// SIMATIC S7-200 project (STEP 7-Micro/WIN), CPU 224 CN REL 02.01

SYMBOL_TABLE USUARIO1
SF               I0.3     // Sensor de objetos
SII              I0.4     // Sensor inductivo (Metal)
SP               I0.5     // Sensor magnetico (plastico)
SM1              I0.7     // Sensor magnetico extendido 1
SM2              I1.0     // Sensor magnetico extendido 2
SM3              I1.1     // Sensor magnetico extendido 3
SB_2             I1.2     // Pulsador de paro
SB_1             I1.3     // Pulsador de marcha
QS               I1.4     // Zeta de emergencia
SA               I1.5     // Selector de modo
Motor            Q0.0     // Motor
KV1              Q0.4     // Cilindro neumatico 1
KV2              Q0.5     // Cilindro neumatico 2
KV3              Q0.6     // Cilindro neumatico 3
HL1              Q0.7     // Piloto indicador de parada
HL2              Q1.0     // Piloto indicador de marcha
HL3              Q1.1     // Piloto indicador de emergencia
E0               M0.0
E1               M0.1
E2               M0.2
E3               M0.3
E4               M0.4
E5               M0.5
E6               M0.6
E7               M0.7
E8               M1.0
E9               M1.1
EP               M1.2
EM               M1.3
END_CTRL         M1.4     // bit de finalizacion del controlador
C_1              VD100
L_k              VD110
r_k              VD120
e_k              VD130
U_k              VD150
Kp               VD160
END_SYMBOL_TABLE

ORGANIZATION_BLOCK PRINCIPAL:OB1
TITLE=COMENTARIOS DEL PROGRAMA
BEGIN
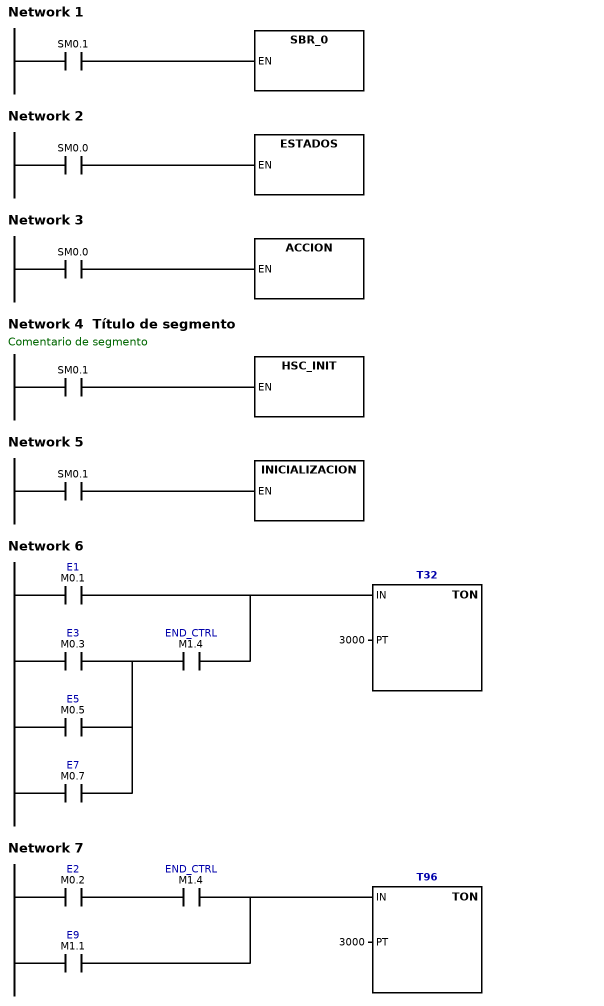
Network 1
LD     SM0.1
CALL   SBR_0:SBR0
Network 2
LD     SM0.0
CALL   ESTADOS:SBR3
Network 3
LD     SM0.0
CALL   ACCION:SBR4
Network 4 // Título de segmento
// Comentario de segmento
LD     SM0.1
CALL   HSC_INIT:SBR1
Network 5
LD     SM0.1
CALL   INICIALIZACION:SBR2
Network 6
LD     E1:M0.1
LD     E3:M0.3
O      E5:M0.5
O      E7:M0.7
A      END_CTRL:M1.4
OLD
TON    T32, 3000
Network 7
LD     E2:M0.2
A      END_CTRL:M1.4
O      E9:M1.1
TON    T96, 3000
END_ORGANIZATION_BLOCK

SUBROUTINE_BLOCK SBR_0:SBR0
TITLE=COMENTARIOS DE LA SUBRUTINA
BEGIN
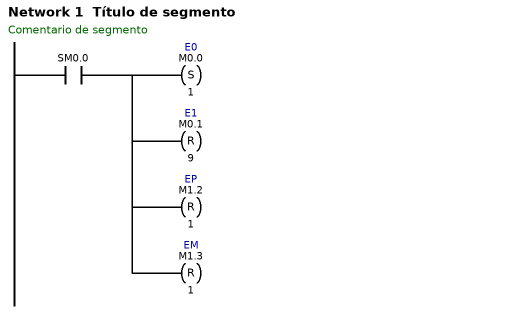
Network 1 // Título de segmento
// Comentario de segmento
LD     SM0.0
S      E0:M0.0, 1
R      E1:M0.1, 9
R      EP:M1.2, 1
R      EM:M1.3, 1
END_SUBROUTINE_BLOCK

SUBROUTINE_BLOCK HSC_INIT:SBR1
TITLE=
BEGIN
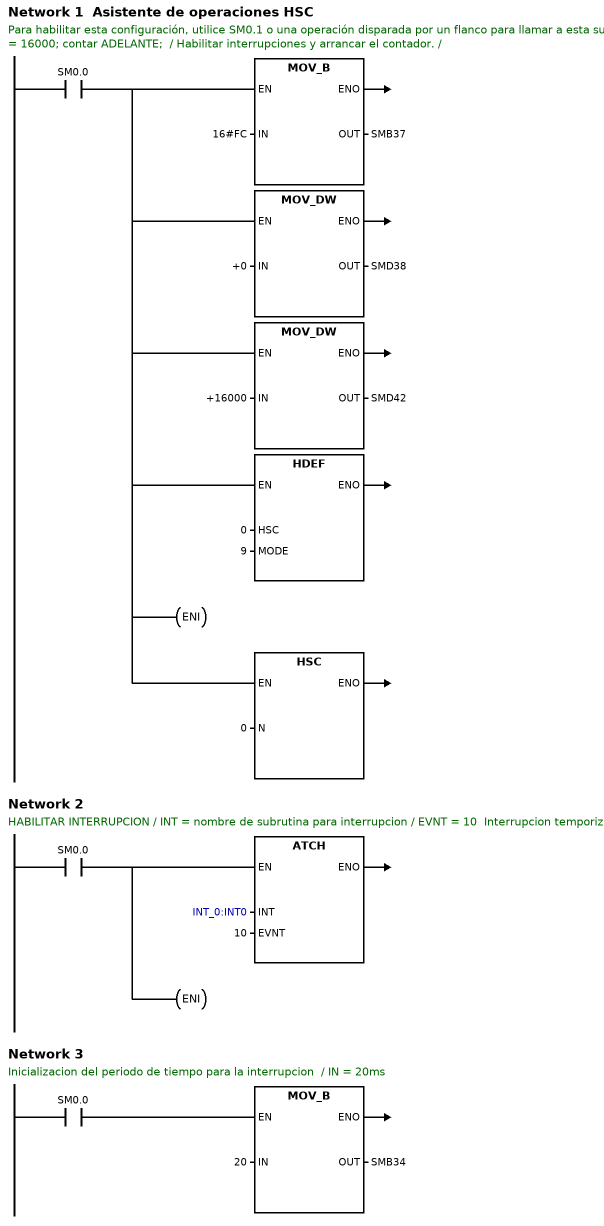
Network 1 // Asistente de operaciones HSC
// Para habilitar esta configuración, utilice SM0.1 o una operación disparada por un flanco para llamar a esta subrutina una vez desde el programa PRINCIPAL. 
// Configurar HC0 para modo 9; CV = 0; PV = 16000; contar ADELANTE; 
// Habilitar interrupciones y arrancar el contador.
// 
//Activar bits de control: contar ADELANTE; velocidad simple; habilitado; 
//Cargar valor actual (CV)
//Cargar valor de preselección (PV)
LD     SM0.0
MOVB   16#FC, SMB37
MOVD   +0, SMD38
MOVD   +16000, SMD42
HDEF   0, 9
ENI
HSC    0
Network 2
// HABILITAR INTERRUPCION
// INT = nombre de subrutina para interrupcion
// EVNT = 10  Interrupcion temporizada 0 SMB34
LD     SM0.0
ATCH   INT_0:INT0, 10
ENI
Network 3
// Inicializacion del periodo de tiempo para la interrupcion 
// IN = 20ms
LD     SM0.0
MOVB   20, SMB34
END_SUBROUTINE_BLOCK

SUBROUTINE_BLOCK INICIALIZACION:SBR2
TITLE=COMENTARIOS DE LA SUBRUTINA
BEGIN
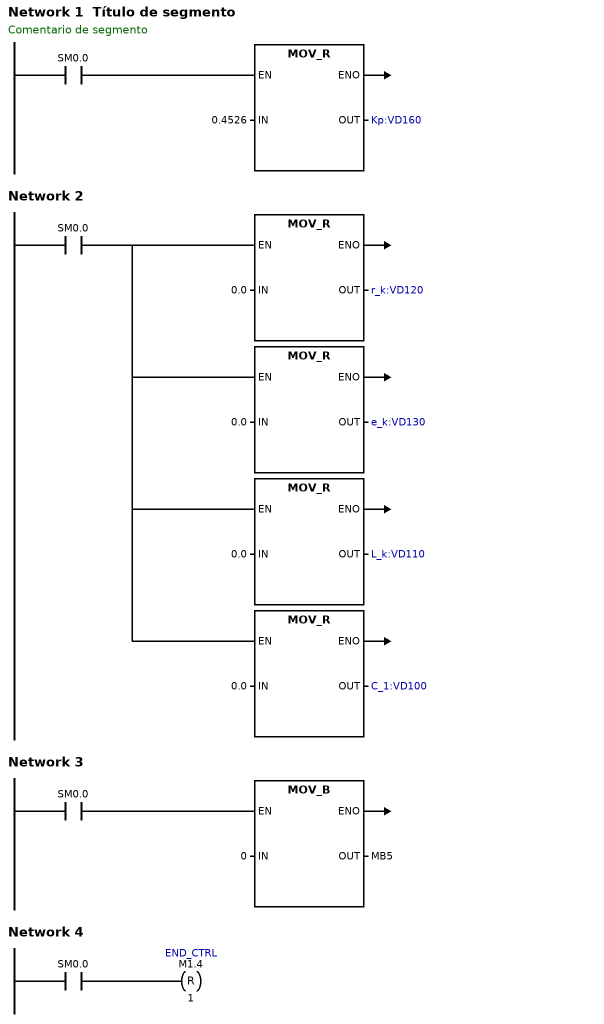
Network 1 // Título de segmento
// Comentario de segmento
LD     SM0.0
MOVR   0.4526, Kp:VD160
Network 2
LD     SM0.0
MOVR   0.0, r_k:VD120
MOVR   0.0, e_k:VD130
MOVR   0.0, L_k:VD110
MOVR   0.0, C_1:VD100
Network 3
LD     SM0.0
MOVB   0, MB5
Network 4
LD     SM0.0
R      END_CTRL:M1.4, 1
END_SUBROUTINE_BLOCK

SUBROUTINE_BLOCK ESTADOS:SBR3
TITLE=COMENTARIOS DE LA SUBRUTINA
BEGIN
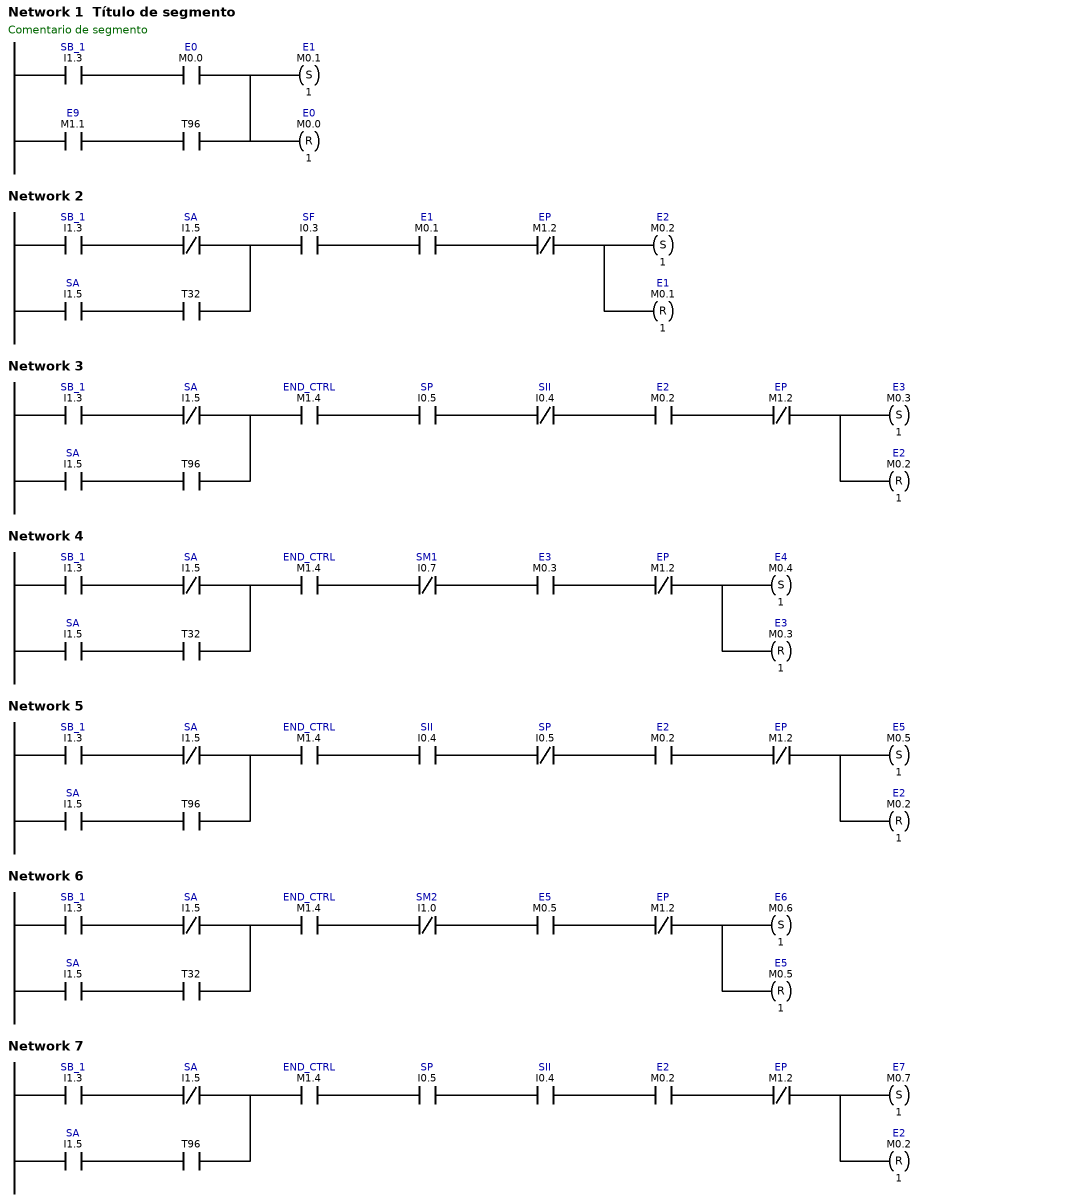
Network 1 // Título de segmento
// Comentario de segmento
LD     SB_1:I1.3
A      E0:M0.0
LD     E9:M1.1
A      T96
OLD
S      E1:M0.1, 1
R      E0:M0.0, 1
Network 2
LD     SB_1:I1.3
AN     SA:I1.5
LD     SA:I1.5
A      T32
OLD
A      SF:I0.3
A      E1:M0.1
AN     EP:M1.2
S      E2:M0.2, 1
R      E1:M0.1, 1
Network 3
LD     SB_1:I1.3
AN     SA:I1.5
LD     SA:I1.5
A      T96
OLD
A      END_CTRL:M1.4
A      SP:I0.5
AN     SII:I0.4
A      E2:M0.2
AN     EP:M1.2
S      E3:M0.3, 1
R      E2:M0.2, 1
Network 4
LD     SB_1:I1.3
AN     SA:I1.5
LD     SA:I1.5
A      T32
OLD
A      END_CTRL:M1.4
AN     SM1:I0.7
A      E3:M0.3
AN     EP:M1.2
S      E4:M0.4, 1
R      E3:M0.3, 1
Network 5
LD     SB_1:I1.3
AN     SA:I1.5
LD     SA:I1.5
A      T96
OLD
A      END_CTRL:M1.4
A      SII:I0.4
AN     SP:I0.5
A      E2:M0.2
AN     EP:M1.2
S      E5:M0.5, 1
R      E2:M0.2, 1
Network 6
LD     SB_1:I1.3
AN     SA:I1.5
LD     SA:I1.5
A      T32
OLD
A      END_CTRL:M1.4
AN     SM2:I1.0
A      E5:M0.5
AN     EP:M1.2
S      E6:M0.6, 1
R      E5:M0.5, 1
Network 7
LD     SB_1:I1.3
AN     SA:I1.5
LD     SA:I1.5
A      T96
OLD
A      END_CTRL:M1.4
A      SP:I0.5
A      SII:I0.4
A      E2:M0.2
AN     EP:M1.2
S      E7:M0.7, 1
R      E2:M0.2, 1
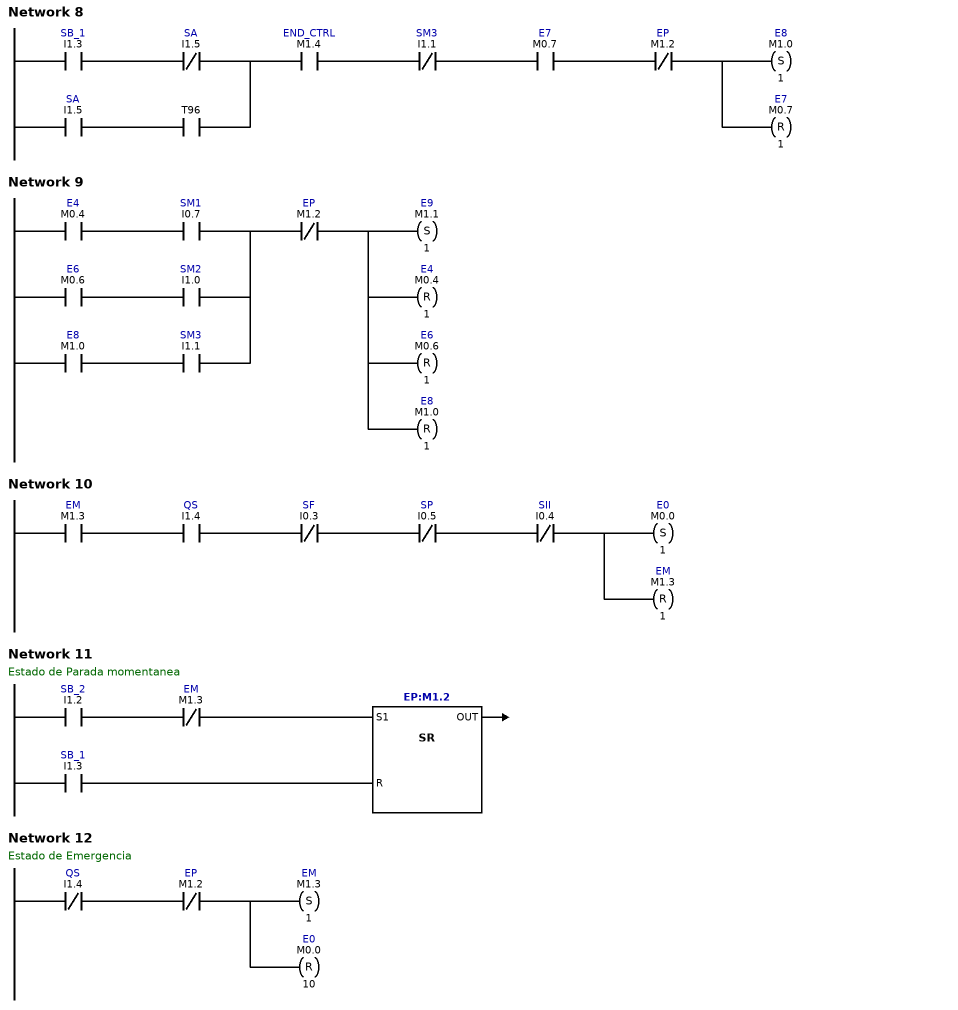
Network 8
LD     SB_1:I1.3
AN     SA:I1.5
LD     SA:I1.5
A      T96
OLD
A      END_CTRL:M1.4
AN     SM3:I1.1
A      E7:M0.7
AN     EP:M1.2
S      E8:M1.0, 1
R      E7:M0.7, 1
Network 9
LD     E4:M0.4
A      SM1:I0.7
LD     E6:M0.6
A      SM2:I1.0
OLD
LD     E8:M1.0
A      SM3:I1.1
OLD
AN     EP:M1.2
S      E9:M1.1, 1
R      E4:M0.4, 1
R      E6:M0.6, 1
R      E8:M1.0, 1
Network 10
LD     EM:M1.3
A      QS:I1.4
AN     SF:I0.3
AN     SP:I0.5
AN     SII:I0.4
S      E0:M0.0, 1
R      EM:M1.3, 1
Network 11
// Estado de Parada momentanea
LD     SB_2:I1.2
AN     EM:M1.3
LD     SB_1:I1.3
NOT
A      EP:M1.2
OLD
=      EP:M1.2
Network 12
// Estado de Emergencia
LDN    QS:I1.4
AN     EP:M1.2
S      EM:M1.3, 1
R      E0:M0.0, 10
END_SUBROUTINE_BLOCK

SUBROUTINE_BLOCK ACCION:SBR4
TITLE=COMENTARIOS DE LA SUBRUTINA
BEGIN
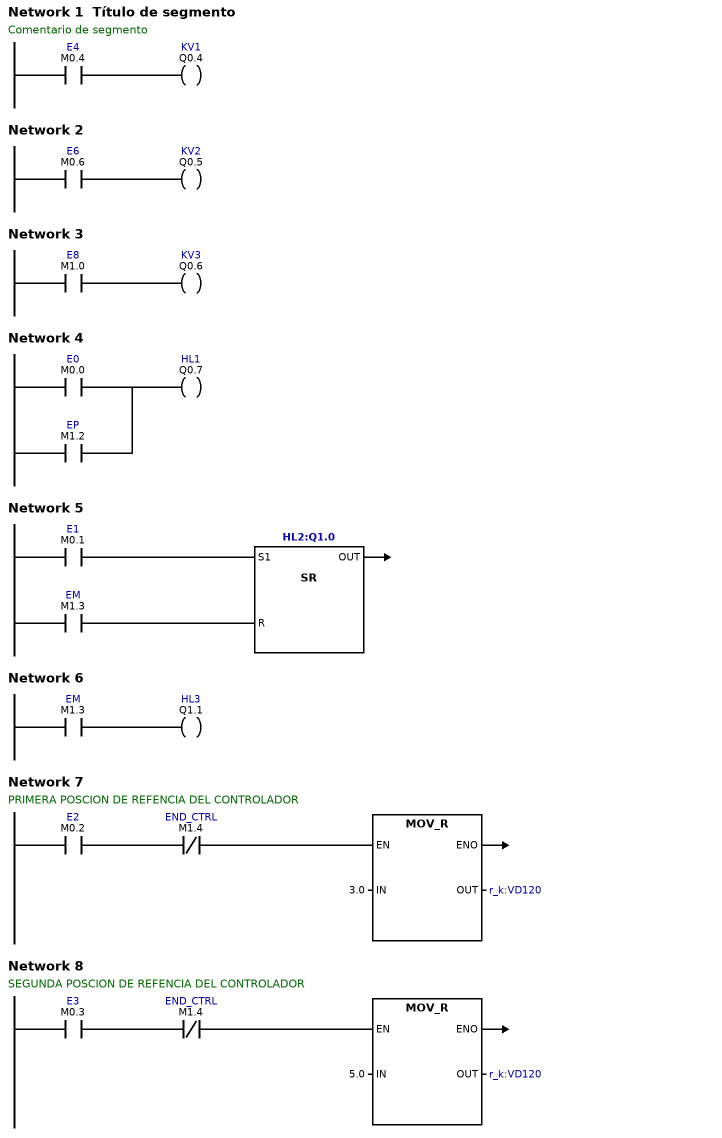
Network 1 // Título de segmento
// Comentario de segmento
LD     E4:M0.4
=      KV1:Q0.4
Network 2
LD     E6:M0.6
=      KV2:Q0.5
Network 3
LD     E8:M1.0
=      KV3:Q0.6
Network 4
LD     E0:M0.0
O      EP:M1.2
=      HL1:Q0.7
Network 5
LD     E1:M0.1
LD     EM:M1.3
NOT
A      HL2:Q1.0
OLD
=      HL2:Q1.0
Network 6
LD     EM:M1.3
=      HL3:Q1.1
Network 7
// PRIMERA POSCION DE REFENCIA DEL CONTROLADOR
LD     E2:M0.2
AN     END_CTRL:M1.4
MOVR   3.0, r_k:VD120
Network 8
// SEGUNDA POSCION DE REFENCIA DEL CONTROLADOR
LD     E3:M0.3
AN     END_CTRL:M1.4
MOVR   5.0, r_k:VD120
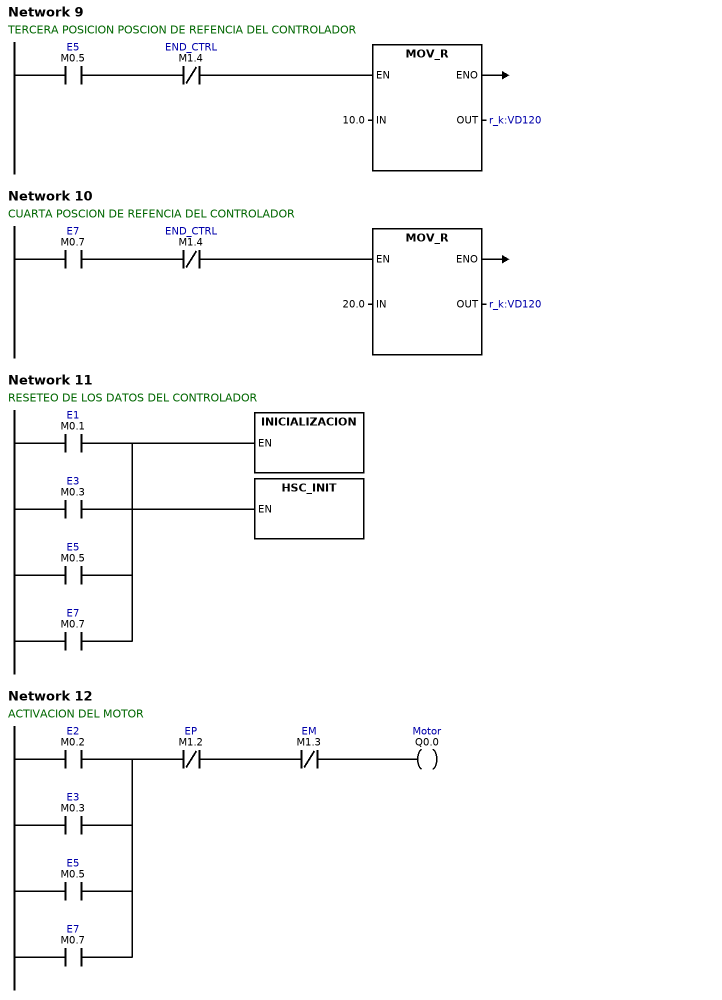
Network 9
// TERCERA POSICION POSCION DE REFENCIA DEL CONTROLADOR
LD     E5:M0.5
AN     END_CTRL:M1.4
MOVR   10.0, r_k:VD120
Network 10
// CUARTA POSCION DE REFENCIA DEL CONTROLADOR
LD     E7:M0.7
AN     END_CTRL:M1.4
MOVR   20.0, r_k:VD120
Network 11
// RESETEO DE LOS DATOS DEL CONTROLADOR
LD     E1:M0.1
O      E3:M0.3
O      E5:M0.5
O      E7:M0.7
CALL   INICIALIZACION:SBR2
CALL   HSC_INIT:SBR1
Network 12
// ACTIVACION DEL MOTOR
LD     E2:M0.2
O      E3:M0.3
O      E5:M0.5
O      E7:M0.7
AN     EP:M1.2
AN     EM:M1.3
=      Motor:Q0.0
END_SUBROUTINE_BLOCK

INTERRUPT_BLOCK INT_0:INT0
TITLE=COMENTARIOS DE LA RUTINA DE INTERRUPCIÓN
BEGIN
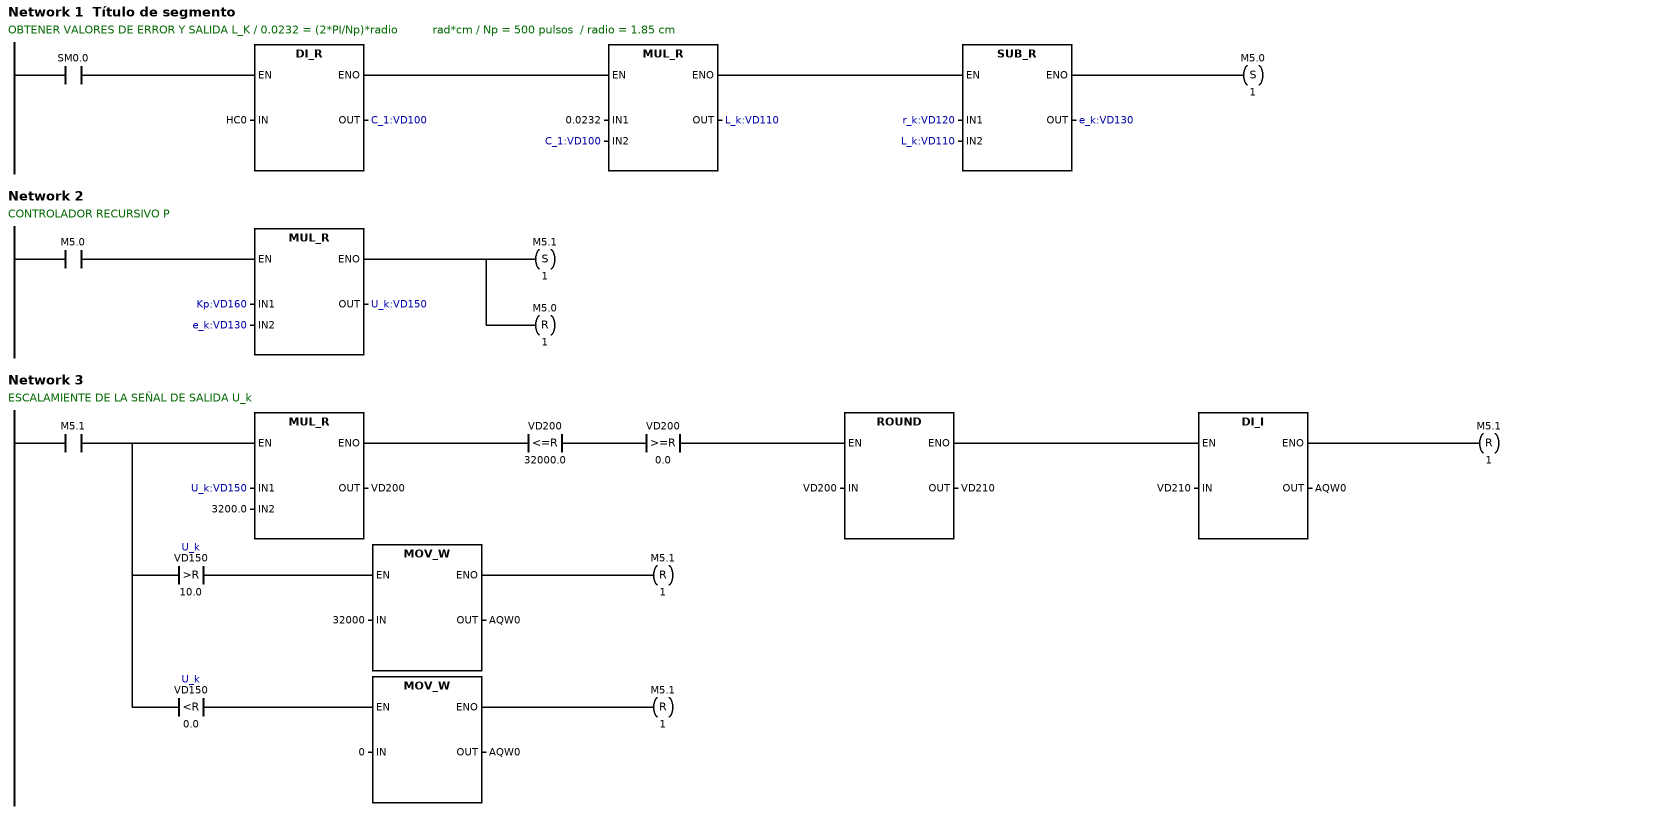
Network 1 // Título de segmento
// OBTENER VALORES DE ERROR Y SALIDA L_K
// 0.0232 = (2*PI/Np)*radio          rad*cm
// Np = 500 pulsos 
// radio = 1.85 cm
LD     SM0.0
DTR    HC0, C_1:VD100
AENO
MOVR   0.0232, L_k:VD110
AENO
*R     C_1:VD100, L_k:VD110
AENO
MOVR   r_k:VD120, e_k:VD130
AENO
-R     L_k:VD110, e_k:VD130
AENO
S      M5.0, 1
Network 2
// CONTROLADOR RECURSIVO P
LD     M5.0
MOVR   Kp:VD160, U_k:VD150
AENO
*R     e_k:VD130, U_k:VD150
AENO
S      M5.1, 1
R      M5.0, 1
Network 3
// ESCALAMIENTE DE LA SEÑAL DE SALIDA U_k
LD     M5.1
LPS
MOVR   U_k:VD150, VD200
AENO
*R     3200.0, VD200
AENO
AR<=   VD200, 32000.0
AR>=   VD200, 0.0
ROUND  VD200, VD210
AENO
DTI    VD210, AQW0
AENO
R      M5.1, 1
LRD
AR>    U_k:VD150, 10.0
MOVW   32000, AQW0
AENO
R      M5.1, 1
LPP
AR<    U_k:VD150, 0.0
MOVW   0, AQW0
AENO
R      M5.1, 1
END_INTERRUPT_BLOCK
